Fanuc KAREL source: KT00239.KL

PROGRAM KT00239
%NOLOCKGROUP
VAR
  I1: INTEGER
  H2: ARRAY[2] OF SHORT
  OUT: BOOLEAN
BEGIN
  I1 = 2
    H2[1] = 3
  OUT = I1 OR H2[1]
END KT00239
